// TIA Portal V21 export
FUNCTION_BLOCK "FB_AnaDoubleAssign"   // FB13, SCL
TITLE = Analyzer: output assigned twice
{ S7_Optimized_Access := 'TRUE' }
// Rule C26e: Motor is assigned twice in one cycle
// stored: MemoryReserve 100, SetENOAutomatically false
   VAR_INPUT
      Start : Bool;   // Start
      Stop : Bool;   // Stop
   END_VAR
   VAR_OUTPUT
      Motor : Bool;   // Motor on
   END_VAR
BEGIN

       #Motor := #Start;
       #Motor := #Motor AND NOT #Stop;
END_FUNCTION_BLOCK
